// Mitsubishi GX Works2 project: PLC_HMI연동   PLC: Q02/Q02H

PROGRAM MAIN
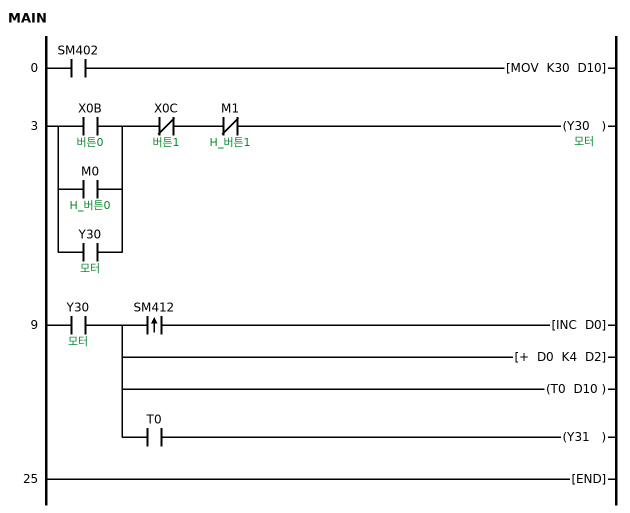
0     LD      SM402
      MOV     K30 D10
3     LD      X0B  ; 버튼0
      OR      M0  ; H_버튼0
      OR      Y30  ; 모터
      ANI     X0C  ; 버튼1
      ANI     M1  ; H_버튼1
      OUT     Y30  ; 모터
9     LD      Y30  ; 모터
      MPS
      ANDP    SM412
      INC     D0
      MPP
      +       D0 K4 D2
      OUT     T0 D10
      AND     T0
      OUT     Y31
25    END
END_PROGRAM

// device comments not shown above
X0  ; 버튼0
X1  ; 버튼1
Y20  ; 모터
